(* IEC 61131-3 sources: Test-Git_ESME26/TestProgettoESME_26.fbsproj/PacDriveLib Migration/Motion/Control/PDL_FB_YOffsetCorrection.fb.st^, 4 files *)

(* ---- ifGetControlChannel.prop.st ---- *)
{attribute 'monitoring' := 'call'}
PROPERTY ifGetControlChannel : MOIN.IF_Axis
__GETTERDECLARATION__
VAR
END_VAR
__GETTERIMPLEMENTATION__

ifGetControlChannel := ifControlChannel;

(* ---- ifGetOffsetChannel.prop.st ---- *)
{attribute 'monitoring' := 'call'}
PROPERTY ifGetOffsetChannel : MOIN.IF_Axis
__GETTERDECLARATION__
VAR
END_VAR
__GETTERIMPLEMENTATION__

ifGetOffsetChannel := ifOffsetChannel;

(* ---- Init.meth.st ---- *)
METHOD PRIVATE Init : BOOL
VAR_INPUT
END_VAR

Init := FALSE;

//check axis
IF i_lencMaster = 0 THEN
	SetDiagOutput(	i_etDiag	:= GD.ET_Diag.InputParameterInvalid,
					i_etDiagExt := PDL_ET_DiagExt.DriveInvalid,
					i_sMsg		:= 'i_lencMaster - Invalid Interface');
	RETURN;

END_IF

Init := TRUE;

(* ---- SetDiagOutput.meth.st ---- *)
{attribute 'hide'}
METHOD SetDiagOutput : BOOL
VAR_INPUT
	i_etDiag	: GD.ET_Diag;
	i_etDiagExt	: PDL_ET_DiagExt;
	i_sMsg		: STRING[80];
END_VAR
VAR
END_VAR

IF i_etDiag <> GD.ET_Diag.Ok THEN
	q_xReady := FALSE;
END_IF

IF q_etDiag = GD.ET_Diag.OK OR i_etDiagExt = PDL_ET_DiagExt.Disabled THEN

	q_etDiag 	:= i_etDiag;
	q_etDiagExt := i_etDiagExt;
	q_sMsg 		:= i_sMsg;

END_IF
